// TIA Portal V18 export
DATA_BLOCK "DB_MB_TCP_ServerConfig"   // DB6
{ S7_Optimized_Access := 'FALSE' }
   VAR RETAIN
      Connect : TCON_IP_v4;
      MB_Disconnect : Bool;
      MB_NDR : Bool;
      MB_DR : Bool;
      MB_Error : Bool;
      MB_Status : Word;
      HoldingReg { S7_SetPoint := 'True'} : Array[0..20] of Word;
   END_VAR
BEGIN
   Connect.InterfaceId := 64;
   Connect.ID := 1;
   Connect.ConnectionType := 11;
   Connect.RemoteAddress.ADDR[1..4] := 0;
   Connect.LocalPort := 502;
   // HoldingReg[0] : MotorOn_Cmd (0=Stop, <>0=Start)
   // HoldingReg[1] : SetFrequency_Hold
   // HoldingReg[2] : FrequencyAct_Hold
   // HoldingReg[3] : MinValueClamp
   // HoldingReg[4] : MaxValueClamp
   // HoldingReg[5] : frequencySource (Выбор источника задания частоты)
END_DATA_BLOCK
